(* IEC 61131-3 sources: bcs-engineering-dsl/language/test/generating/when_test/expected, 2 files *)

(* ---- MAIN_decl.st ---- *)
PROGRAM MAIN
VAR
    x: INT;
    y: BOOL;
    R_TRIG_UnitInstance_ScheduledUnit1: R_TRIG;
    R_TRIG_UnitInstance_OnceConditionalUnit2: R_TRIG;
    fbLocalTime: FB_LocalSystemTime := (bEnable := TRUE);
    timeNow: TIMESTRUCT;
    todNow: TIME_OF_DAY;
    dNow: DATE;
END_VAR

(* ---- MAIN_impl.st ---- *)
fbLocalTime();
timeNow := fbLocalTime.systemTime;
todNow := SYSTEMTIME_TO_TOD(timeNow);
dNow := DT_TO_DATE(SYSTEMTIME_TO_DT(timeNow));

// Scheduled Control Unit 'ScheduledUnit' @ TOD#08:00:00
R_TRIG_UnitInstance_ScheduledUnit1(CLK := todNow >= TOD#08:00:00);
IF R_TRIG_UnitInstance_ScheduledUnit1.Q THEN
    x := 1;
END_IF;

// Conditional Control Unit 'ConditionalUnit'
IF x > 0 THEN
    y := TRUE;
END_IF;

// Conditional Control Unit 'OnceConditionalUnit' (runOnce)
R_TRIG_UnitInstance_OnceConditionalUnit2(CLK := y);
IF R_TRIG_UnitInstance_OnceConditionalUnit2.Q THEN
    x := 2;
END_IF;
